{region 'Documentation'}
(*!
<summary>Checks that unused array capacity at indices 4 through 6 is never processed.</summary>
*)
{endregion}
FUNCTION_BLOCK Test_OrchestratorUnusedCapacity EXTENDS OrchestrationTestBase

SUPER^();

{region 'Documentation'}
(*!
<summary>Defines this scenario independently of the subject's internal fields.</summary>
*)
{endregion}
METHOD PROTECTED ConfigureScenario
FArrayLayout := E_OrchestrationArrayLayout.SpareCapacity;
FChildCount := 3;
ConfigureStandardSequence();
END_METHOD

END_FUNCTION_BLOCK

(* stored: Version 1.1.0.1
   POU Test_OrchestratorUnusedCapacity: Id {862839a5-5ded-4ccc-8b4b-7048c19cde23}, SpecialFunc None
   Folder Internal: Id {4562e2ef-b109-4664-aad7-297cb79cd611}
   Method ConfigureScenario: Id {dfd7b03a-1bf4-459e-9c4d-1f0def2dd489} *)
